(* INIT DIGITAL OUTPUT STUFF *)
FB_DO_SW_001.InitMqtt(MQTTPublishPrefix:= ADR(MqttPubSwitchPrefix),					(* pointer to string prefix for the mqtt publish topic *)
	MQTTSubscribePrefix:= ADR(MqttSubSwitchPrefix),									(* pointer to string prefix for the mqtt subscribe topic *)
	pMqttPublishQueue := ADR(MqttVariables.fbMqttPublishQueue),						(* pointer to MqttPublishQueue to send a new Mqtt event *)
	pMqttCallbackCollector := ADR(MqttVariables.collector_FB_OUTPUT_SWITCH_MQTT)	(* pointer to CallbackCollector to receive Mqtt subscription events *)
);
FB_DO_SW_002.InitMqtt(MQTTPublishPrefix:= ADR(MqttPubSwitchPrefix),	MQTTSubscribePrefix:= ADR(MqttSubSwitchPrefix), pMqttPublishQueue := ADR(MqttVariables.fbMqttPublishQueue), pMqttCallbackCollector := ADR(MqttVariables.collector_FB_OUTPUT_SWITCH_MQTT));
FB_DO_SW_003.InitMqtt(MQTTPublishPrefix:= ADR(MqttPubSwitchPrefix),	MQTTSubscribePrefix:= ADR(MqttSubSwitchPrefix),	pMqttPublishQueue := ADR(MqttVariables.fbMqttPublishQueue), pMqttCallbackCollector := ADR(MqttVariables.collector_FB_OUTPUT_SWITCH_MQTT));
FB_DO_SW_004.InitMqtt(MQTTPublishPrefix:= ADR(MqttPubSwitchPrefix),	MQTTSubscribePrefix:= ADR(MqttSubSwitchPrefix),	pMqttPublishQueue := ADR(MqttVariables.fbMqttPublishQueue), pMqttCallbackCollector := ADR(MqttVariables.collector_FB_OUTPUT_SWITCH_MQTT));
FB_DO_SW_005.InitMqtt(MQTTPublishPrefix:= ADR(MqttPubSwitchPrefix),	MQTTSubscribePrefix:= ADR(MqttSubSwitchPrefix),	pMqttPublishQueue := ADR(MqttVariables.fbMqttPublishQueue), pMqttCallbackCollector := ADR(MqttVariables.collector_FB_OUTPUT_SWITCH_MQTT));
FB_DO_SW_006.InitMqtt(MQTTPublishPrefix:= ADR(MqttPubSwitchPrefix),	MQTTSubscribePrefix:= ADR(MqttSubSwitchPrefix),	pMqttPublishQueue := ADR(MqttVariables.fbMqttPublishQueue), pMqttCallbackCollector := ADR(MqttVariables.collector_FB_OUTPUT_SWITCH_MQTT));
FB_DO_SW_007.InitMqtt(MQTTPublishPrefix:= ADR(MqttPubSwitchPrefix),	MQTTSubscribePrefix:= ADR(MqttSubSwitchPrefix),	pMqttPublishQueue := ADR(MqttVariables.fbMqttPublishQueue), pMqttCallbackCollector := ADR(MqttVariables.collector_FB_OUTPUT_SWITCH_MQTT));
FB_DO_SW_008.InitMqtt(MQTTPublishPrefix:= ADR(MqttPubSwitchPrefix),	MQTTSubscribePrefix:= ADR(MqttSubSwitchPrefix),	pMqttPublishQueue := ADR(MqttVariables.fbMqttPublishQueue), pMqttCallbackCollector := ADR(MqttVariables.collector_FB_OUTPUT_SWITCH_MQTT));
FB_DO_SW_009.InitMqtt(MQTTPublishPrefix:= ADR(MqttPubSwitchPrefix),	MQTTSubscribePrefix:= ADR(MqttSubSwitchPrefix),	pMqttPublishQueue := ADR(MqttVariables.fbMqttPublishQueue), pMqttCallbackCollector := ADR(MqttVariables.collector_FB_OUTPUT_SWITCH_MQTT));
FB_DO_SW_010.InitMqtt(MQTTPublishPrefix:= ADR(MqttPubSwitchPrefix),	MQTTSubscribePrefix:= ADR(MqttSubSwitchPrefix),	pMqttPublishQueue := ADR(MqttVariables.fbMqttPublishQueue), pMqttCallbackCollector := ADR(MqttVariables.collector_FB_OUTPUT_SWITCH_MQTT));
FB_DO_SW_011.InitMqtt(MQTTPublishPrefix:= ADR(MqttPubSwitchPrefix),	MQTTSubscribePrefix:= ADR(MqttSubSwitchPrefix),	pMqttPublishQueue := ADR(MqttVariables.fbMqttPublishQueue), pMqttCallbackCollector := ADR(MqttVariables.collector_FB_OUTPUT_SWITCH_MQTT));
FB_DO_SW_012.InitMqtt(MQTTPublishPrefix:= ADR(MqttPubSwitchPrefix),	MQTTSubscribePrefix:= ADR(MqttSubSwitchPrefix), pMqttPublishQueue := ADR(MqttVariables.fbMqttPublishQueue), pMqttCallbackCollector := ADR(MqttVariables.collector_FB_OUTPUT_SWITCH_MQTT));
FB_DO_SW_013.InitMqtt(MQTTPublishPrefix:= ADR(MqttPubSwitchPrefix),	MQTTSubscribePrefix:= ADR(MqttSubSwitchPrefix), pMqttPublishQueue := ADR(MqttVariables.fbMqttPublishQueue), pMqttCallbackCollector := ADR(MqttVariables.collector_FB_OUTPUT_SWITCH_MQTT));
FB_DO_SW_014.InitMqtt(MQTTPublishPrefix:= ADR(MqttPubSwitchPrefix),	MQTTSubscribePrefix:= ADR(MqttSubSwitchPrefix), pMqttPublishQueue := ADR(MqttVariables.fbMqttPublishQueue), pMqttCallbackCollector := ADR(MqttVariables.collector_FB_OUTPUT_SWITCH_MQTT));
FB_DO_SW_015.InitMqtt(MQTTPublishPrefix:= ADR(MqttPubSwitchPrefix),	MQTTSubscribePrefix:= ADR(MqttSubSwitchPrefix), pMqttPublishQueue := ADR(MqttVariables.fbMqttPublishQueue), pMqttCallbackCollector := ADR(MqttVariables.collector_FB_OUTPUT_SWITCH_MQTT));
FB_DO_SW_016.InitMqtt(MQTTPublishPrefix:= ADR(MqttPubSwitchPrefix),	MQTTSubscribePrefix:= ADR(MqttSubSwitchPrefix), pMqttPublishQueue := ADR(MqttVariables.fbMqttPublishQueue), pMqttCallbackCollector := ADR(MqttVariables.collector_FB_OUTPUT_SWITCH_MQTT));
FB_DO_SW_017.InitMqtt(MQTTPublishPrefix:= ADR(MqttPubSwitchPrefix),	MQTTSubscribePrefix:= ADR(MqttSubSwitchPrefix), pMqttPublishQueue := ADR(MqttVariables.fbMqttPublishQueue), pMqttCallbackCollector := ADR(MqttVariables.collector_FB_OUTPUT_SWITCH_MQTT));
FB_DO_SW_018.InitMqtt(MQTTPublishPrefix:= ADR(MqttPubSwitchPrefix),	MQTTSubscribePrefix:= ADR(MqttSubSwitchPrefix), pMqttPublishQueue := ADR(MqttVariables.fbMqttPublishQueue), pMqttCallbackCollector := ADR(MqttVariables.collector_FB_OUTPUT_SWITCH_MQTT));
FB_DO_SW_019.InitMqtt(MQTTPublishPrefix:= ADR(MqttPubSwitchPrefix),	MQTTSubscribePrefix:= ADR(MqttSubSwitchPrefix), pMqttPublishQueue := ADR(MqttVariables.fbMqttPublishQueue), pMqttCallbackCollector := ADR(MqttVariables.collector_FB_OUTPUT_SWITCH_MQTT));
FB_DO_SW_020.InitMqtt(MQTTPublishPrefix:= ADR(MqttPubSwitchPrefix),	MQTTSubscribePrefix:= ADR(MqttSubSwitchPrefix), pMqttPublishQueue := ADR(MqttVariables.fbMqttPublishQueue), pMqttCallbackCollector := ADR(MqttVariables.collector_FB_OUTPUT_SWITCH_MQTT));
FB_DO_SW_021.InitMqtt(MQTTPublishPrefix:= ADR(MqttPubSwitchPrefix),	MQTTSubscribePrefix:= ADR(MqttSubSwitchPrefix), pMqttPublishQueue := ADR(MqttVariables.fbMqttPublishQueue), pMqttCallbackCollector := ADR(MqttVariables.collector_FB_OUTPUT_SWITCH_MQTT));
FB_DO_SW_022.InitMqtt(MQTTPublishPrefix:= ADR(MqttPubSwitchPrefix),	MQTTSubscribePrefix:= ADR(MqttSubSwitchPrefix), pMqttPublishQueue := ADR(MqttVariables.fbMqttPublishQueue), pMqttCallbackCollector := ADR(MqttVariables.collector_FB_OUTPUT_SWITCH_MQTT));
FB_DO_SW_023.InitMqtt(MQTTPublishPrefix:= ADR(MqttPubSwitchPrefix),	MQTTSubscribePrefix:= ADR(MqttSubSwitchPrefix), pMqttPublishQueue := ADR(MqttVariables.fbMqttPublishQueue), pMqttCallbackCollector := ADR(MqttVariables.collector_FB_OUTPUT_SWITCH_MQTT));
FB_DO_SW_024.InitMqtt(MQTTPublishPrefix:= ADR(MqttPubSwitchPrefix),	MQTTSubscribePrefix:= ADR(MqttSubSwitchPrefix), pMqttPublishQueue := ADR(MqttVariables.fbMqttPublishQueue), pMqttCallbackCollector := ADR(MqttVariables.collector_FB_OUTPUT_SWITCH_MQTT));
FB_DO_SW_025.InitMqtt(MQTTPublishPrefix:= ADR(MqttPubSwitchPrefix),	MQTTSubscribePrefix:= ADR(MqttSubSwitchPrefix), pMqttPublishQueue := ADR(MqttVariables.fbMqttPublishQueue), pMqttCallbackCollector := ADR(MqttVariables.collector_FB_OUTPUT_SWITCH_MQTT));
FB_DO_SW_026.InitMqtt(MQTTPublishPrefix:= ADR(MqttPubSwitchPrefix),	MQTTSubscribePrefix:= ADR(MqttSubSwitchPrefix), pMqttPublishQueue := ADR(MqttVariables.fbMqttPublishQueue), pMqttCallbackCollector := ADR(MqttVariables.collector_FB_OUTPUT_SWITCH_MQTT));
FB_DO_SW_027.InitMqtt(MQTTPublishPrefix:= ADR(MqttPubSwitchPrefix),	MQTTSubscribePrefix:= ADR(MqttSubSwitchPrefix), pMqttPublishQueue := ADR(MqttVariables.fbMqttPublishQueue), pMqttCallbackCollector := ADR(MqttVariables.collector_FB_OUTPUT_SWITCH_MQTT));
FB_DO_SW_028.InitMqtt(MQTTPublishPrefix:= ADR(MqttPubSwitchPrefix),	MQTTSubscribePrefix:= ADR(MqttSubSwitchPrefix), pMqttPublishQueue := ADR(MqttVariables.fbMqttPublishQueue), pMqttCallbackCollector := ADR(MqttVariables.collector_FB_OUTPUT_SWITCH_MQTT));
FB_DO_SW_029.InitMqtt(MQTTPublishPrefix:= ADR(MqttPubSwitchPrefix),	MQTTSubscribePrefix:= ADR(MqttSubSwitchPrefix), pMqttPublishQueue := ADR(MqttVariables.fbMqttPublishQueue), pMqttCallbackCollector := ADR(MqttVariables.collector_FB_OUTPUT_SWITCH_MQTT));
FB_DO_SW_030.InitMqtt(MQTTPublishPrefix:= ADR(MqttPubSwitchPrefix),	MQTTSubscribePrefix:= ADR(MqttSubSwitchPrefix), pMqttPublishQueue := ADR(MqttVariables.fbMqttPublishQueue), pMqttCallbackCollector := ADR(MqttVariables.collector_FB_OUTPUT_SWITCH_MQTT));

(* INIT COVERS STUFF *)
FB_DO_COVER_001.InitMqtt(MQTTPublishPrefix:= ADR(MqttPubCoverPrefix),				(* pointer to string prefix for the mqtt publish topic *)
	MQTTSubscribePrefix:= ADR(MqttSubCoverPrefix),									(* pointer to string prefix for the mqtt subscribe topic *)
	pMqttPublishQueue := ADR(MqttVariables.fbMqttPublishQueue),						(* pointer to MqttPublishQueue to send a new Mqtt event *)
	pMqttCallbackCollector := ADR(MqttVariables.collector_FB_OUTPUT_COVER_MQTT), 	(* pointer to CallbackCollector to receive Mqtt subscription events *)
	MQTT.QoS.ExactlyOnce, 														(* specify the QoS for the POS mqtt events (values 0-100) *)
	2																				(* specify the resolution for the POS mqtt events *)
);

FB_DO_COVER_001.ConfigureFunctionBlock(T_LOCKOUT:=T#1S,								(* delay between change of direction *)
	T_UD:=T#20S																		(* run time to move the cover completely up/down *)
);

(* INIT VIRTUAL STUFF *)
FB_VIRTUAL_STRING_001.InitMqtt(MQTTPublishPrefix:= ADR(MqttPubVirtualPrefix),				
	MQTTSubscribePrefix:= ADR(MqttSubVirtualPrefix),									
	pMqttPublishQueue := ADR(MqttVariables.fbMqttPublishQueue),						
	pMqttCallbackCollector := ADR(MqttVariables.collector_FB_VIRTUAL_MQTT),
	MqttQos:=MQTT.QoS.ExactlyOnce, 
	MqttRetain:=FALSE									
);
FB_VIRTUAL_STRING_001.ConfigureFunctionBlockAsVirtualInput(DefaultValue:='HelloWorld',SetDefaultValueStartup:=TRUE,PublishAtStartup:=TRUE,UsePersistentAtStartup:=FALSE,ConfirmReceival:=TRUE);


FB_VIRTUAL_INT_001.InitMqtt(MQTTPublishPrefix:= ADR(MqttPubVirtualPrefix),				
	MQTTSubscribePrefix:= ADR(MqttSubVirtualPrefix),									
	pMqttPublishQueue := ADR(MqttVariables.fbMqttPublishQueue),						
	pMqttCallbackCollector := ADR(MqttVariables.collector_FB_VIRTUAL_MQTT),
	MqttQos:=MQTT.QoS.ExactlyOnce, 
	MqttRetain:=FALSE												
);
FB_VIRTUAL_INT_001.ConfigureFunctionBlockAsVirtualInput(DefaultValue:=0,SetDefaultValueStartup:=TRUE,PublishAtStartup:=TRUE,UsePersistentAtStartup:=FALSE,ConfirmReceival:=TRUE);
(* FB_VIRTUAL_INT_001.ConfigureFunctionBlockAsVirtualOutput(PublishAtStartup:=TRUE); *)


FB_VIRTUAL_BOOL_001.InitMqtt(MQTTPublishPrefix:= ADR(MqttPubVirtualPrefix),				
	MQTTSubscribePrefix:= ADR(MqttSubVirtualPrefix),									
	pMqttPublishQueue := ADR(MqttVariables.fbMqttPublishQueue),						
	pMqttCallbackCollector := ADR(MqttVariables.collector_FB_VIRTUAL_MQTT),
	MqttQos:=MQTT.QoS.ExactlyOnce, 
	MqttRetain:=FALSE											
);
(* FB_VIRTUAL_BOOL_001.ConfigureFunctionBlockAsVirtualInput(DefaultValue:=FALSE,SetDefaultValueStartup:=TRUE,PublishAtStartup:=TRUE,UsePersistentAtStartup:=FALSE); *)
FB_VIRTUAL_BOOL_001.ConfigureFunctionBlockAsVirtualOutput(PublishAtStartup:=TRUE);

FB_VIRTUAL_REAL_001.InitMqtt(MQTTPublishPrefix:= ADR(MqttPubVirtualPrefix),				
	MQTTSubscribePrefix:= ADR(MqttSubVirtualPrefix),									
	pMqttPublishQueue := ADR(MqttVariables.fbMqttPublishQueue),						
	pMqttCallbackCollector := ADR(MqttVariables.collector_FB_VIRTUAL_MQTT),
	MqttQos:=MQTT.QoS.ExactlyOnce, 
	MqttRetain:=FALSE												
);
FB_VIRTUAL_REAL_001.ConfigureFunctionBlockAsVirtualInput(DefaultValue:=0.1,SetDefaultValueStartup:=TRUE,PublishAtStartup:=TRUE,UsePersistentAtStartup:=FALSE,ConfirmReceival:=TRUE);
(* FB_VIRTUAL_REAL_001.ConfigureFunctionBlockAsVirtualOutput(PublishAtStartup:=TRUE); *)


(* INIT BISTABLE RELAIS *) 
FB_DO_BISTABLE_001.InitMqtt(MQTTPublishPrefix:= ADR(MqttPubSwitchPrefix),	MQTTSubscribePrefix:= ADR(MqttSubSwitchPrefix), pMqttPublishQueue := ADR(MqttVariables.fbMqttPublishQueue), pMqttCallbackCollector := ADR(MqttVariables.collector_FB_OUTPUT_SWITCH_MQTT));
FB_DO_BISTABLE_001.ConfigureFunctionBlock(T_hold:=T#10S); 

                    
END_ACTION

ACTION MOVE_COVERS:
                      FB_DO_COVER_001(
	UP:=FB_DI_PB_013.P_LONG,
	DN:=FB_DI_PB_015.P_LONG,
	MU=>DO_031,
	MD=>DO_032	
	);
                    
END_ACTION

ACTION PROCESS_VIRTUAL:
                      
FB_VIRTUAL_BOOL_001();
FB_VIRTUAL_INT_001();
FB_VIRTUAL_STRING_001();
FB_VIRTUAL_REAL_001();
                    
END_ACTION
END_PROGRAM

PROGRAM PLC_PRG_MQTT
  VAR
    broker : STRING := '192.168.1.52:1883';  (* variables for MQTT configuration *)
    clientID : STRING := 'PLC-House';  (* use the below for username password authentication to broker broker :STRING:='user:password@192.168.1.36:1883'; user led to indicate broker status, é!COCKPIT version LED_1_BrokerStatus :FbAppLED; *)
    MQTTClient : MQTT.MQTTClient;
    MQTT_IN_OUT : MQTT.MQTT_IN_OUT;
    MQTTInfo : MQTT.MQTT_INFO;
    MQTTLwtTopic : STRING := 'Devices/PLC/House/availability';
    MQTTLwtPayload : STRING := 'offline';
    MQTTBirthMessage : MQTT_MESSAGE;
    MQTTBirthTopic : STRING := 'Devices/PLC/House/availability';
    MQTTBirthPayload : STRING := 'online';
    MQTTBirthHartbeat : OSCAT_BASIC.GEN_PULSE;
    MQTTBirthHartbeatTime : TIME := TIME#5s0ms;
    MQTTConnectTrigger : Standard.R_TRIG;
    MQTTPublishBirth : BOOL := TRUE;
    MQTTBirthPublisher : FB_MqttPublishWorker;
    initMqtt : BOOL;  (* variables for MQTT setup *)
    icounter : UDINT;
    ipublishers : UDINT := 40;  (* variables for MQTT publishing *)
    publishers : ARRAY[0..39] OF FB_MqttPublishWorker;
    i : UDINT;  (* variables to work with Mqttbuffer *)
    subscriber_FB_OUTPUT_SWITCH_MQTT : MQTT.MQTTSubscribe;  (* variables for MQTT subscribing *)
    subscriber_FB_OUTPUT_COVER_MQTT : MQTT.MQTTSubscribe;
    subscriber_FB_VIRTUAL_MQTT : MQTT.MQTTSubscribe;
    subscriber_FB_DIMMER_MQTT : MQTT.MQTTSubscribe;
  END_VAR

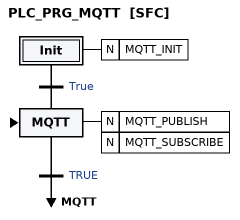
INITIAL_STEP Init:
  MQTT_INIT(N);
END_STEP
TRANSITION FROM Init TO MQTT
  := True;
END_TRANSITION
STEP MQTT:
  MQTT_PUBLISH(N);
  MQTT_SUBSCRIBE(N);
END_STEP
TRANSITION FROM MQTT TO MQTT
  := TRUE;
END_TRANSITION

ACTION MQTT_INIT:
                      
IF NOT initMqtt THEN
	initMqtt := TRUE;
	(* Basic MQTT config *)
	MQTT_IN_OUT.ClientID := clientID;
	
	(* Set the LWT topic / payload *)
	MQTT_IN_OUT.BuildWillTopicAndMessage := FALSE;
	MQTT_IN_OUT.WillTopicBase := '';
	MQTT_IN_OUT.ClientWillTopic := MQTTLwtTopic;
	MQTT_IN_OUT.ClientWillMessage := MQTTLwtPayload;
	
	(* Set the birth message *)
	MQTTBirthMessage.Payload := MQTTBirthPayload;
	MQTTBirthMessage.Topic := MQTTBirthTopic;
	MQTTBirthMessage.Qos := MqttVariables.MQTT_QOS_EXACTLY_ONCE;
	MQTTBirthMessage.MqttRetain := FALSE;
	
	(* Configure the rising edge detector to detect a connect/reconnect to the broker, used for  birth message *)
	MQTTConnectTrigger(CLK := MQTTInfo.MQTT_CONNECTED);
	
	(* Configure the dedicated MQTTBirth publisher *)
	MQTTBirthPublisher.Init(inputMQTT_IN_OUT:= ADR(MQTT_IN_OUT));
	
	(* Configure the pulse generator for the birth message hartbeat *)
	 MQTTBirthHartbeat(ENQ:=TRUE, PTH:=T#0S, PTL:=MQTTBirthHartbeatTime);
	
	(* INIT MQTT PUBLISH STUFF *)
	FOR icounter := 0 TO (ipublishers-1) DO		
		publishers[icounter].Init(inputMQTT_IN_OUT:= ADR(MQTT_IN_OUT));
	END_FOR 
	
	(* INIT MQTT SUBSCRIBE STUFF *)
	subscriber_FB_OUTPUT_SWITCH_MQTT.SetMqttInOut(MQTT_IN_OUT:= MQTT_IN_OUT);	
	subscriber_FB_OUTPUT_COVER_MQTT.SetMqttInOut(MQTT_IN_OUT:= MQTT_IN_OUT);
	subscriber_FB_VIRTUAL_MQTT.SetMqttInOut(MQTT_IN_OUT:= MQTT_IN_OUT);	
	subscriber_FB_DIMMER_MQTT.SetMqttInOut(MQTT_IN_OUT:= MQTT_IN_OUT);

END_IF


                    
END_ACTION

ACTION MQTT_PUBLISH:
                      (* set user led green if connected to MQTT broker, flashing red if not *)
(* é!COCKPIT version *)
(* LED_1_BrokerStatus(eID:=eLedID.AppLED_1, xOpen:=TRUE );
IF(MQTTClient.connected) THEN
	LED_1_BrokerStatus.SetStatic(eLedColor.Green);
ELSE
	LED_1_BrokerStatus.SetFlash(T#1S,eLedColor.Red, eLedColor.Off);  
END_IF *)
(* Codesys 3S version *)
(*
IF MQTTClient.connected THEN
     PFC.SetLed(which:=PFC.LED.U1, how:=PFC.LedState.STATIC_GRN);
ELSE
     PFC.SetLed(which:=PFC.LED.U1, how:=PFC.LedState.BLINK_RED);
END_IF 
*)

(* allow the rising edge detector to detect a connect/reconnect to the broker, used for  birth message *)
MQTTConnectTrigger(CLK := MQTTInfo.MQTT_CONNECTED);

(* allow the pulse generator to generate a pulse, used for birth message hartbeat *)
MQTTBirthHartbeat(ENQ:=TRUE, PTH:=T#0S, PTL:=MQTTBirthHartbeatTime);

(* Check if this is a new connection due to startup or connection issues *)
IF initMqtt AND (MQTTConnectTrigger.Q OR MQTTBirthHartbeat.Q) THEN
	MQTTPublishBirth := TRUE;
END_IF

(* On connect or reconnect publish a birth message using the dedicated birth publisher *)
IF MQTTPublishBirth THEN
	MQTTBirthPublisher.PublishMessage(MqttMessage := MQTTBirthMessage);
	MQTTPublishBirth:=FALSE;
END_IF


(* Check if Mqtt is initialized AND if there are elements on the queue to process AND if a MQTTbirthmessage has been published successfully *)
IF initMqtt AND NOT(MqttVariables.fbMqttPublishQueue.EMPTY) AND MQTTPublishBirth = FALSE AND MQTTBirthPublisher.SendDone THEN	
	(* Loop through all free publishers untill there are no more elements in the queue or no more free publishers *)
	FOR i:=0 TO (ipublishers-1) DO			
		(* use the publishers that are free  *)
		IF publishers[i].SendDone AND NOT(MqttVariables.fbMqttPublishQueue.EMPTY) THEN	
			(* Pass message from the queue to a publisher *)
			publishers[i].PublishMessage(MqttMessage:= MqttVariables.fbMqttPublishQueue.GetMessage());
		ELSIF MqttVariables.fbMqttPublishQueue.EMPTY THEN
			(* Queue is empty, jump out of the for loop	*)
			EXIT;	
		END_IF
	END_FOR
END_IF


(* If MQTT is initialized, let the MqttPublishWorkers do their work *)
IF initMqtt THEN	
	MQTT_IN_OUT.clientFB(
		MQTT_IN_OUT:= MQTT_IN_OUT, 
		ENABLE:= TRUE, 
		URL:= broker, 
		TIMEOUT:= T#1S, 
		TLS:= FALSE);		
		
	MQTTBirthPublisher();
	
	FOR i := 0 TO (ipublishers-1) DO
  		publishers[i]();
	END_FOR

END_IF

                    
END_ACTION

ACTION MQTT_SUBSCRIBE:
                      (* If MQTT is initialized, let the subscriber(s) do its work *)
IF initMqtt THEN
	
	MQTT_IN_OUT.clientFB(
		MQTT_IN_OUT:= MQTT_IN_OUT, 
		ENABLE:= TRUE, 
		URL:= broker, 
		TIMEOUT:= T#1S, 
		TLS:= FALSE);

	subscriber_FB_OUTPUT_SWITCH_MQTT(
		Subscribe:= TRUE, 
		Topic:= ADR('Devices/PLC/House/In/DigitalOutputs/+'), 
		QoSSubscribe:= MqttVariables.MQTT_QOS_EXACTLY_ONCE, 
		ExpectingString:= TRUE, 
		Callback:= MqttVariables.collector_FB_OUTPUT_SWITCH_MQTT,
	);
	
	subscriber_FB_OUTPUT_COVER_MQTT(
		Subscribe:= TRUE, 
		Topic:= ADR('Devices/PLC/House/In/Covers/+'), 
		QoSSubscribe:= MqttVariables.MQTT_QOS_EXACTLY_ONCE, 
		ExpectingString:= TRUE, 
		Callback:= MqttVariables.collector_FB_OUTPUT_COVER_MQTT,
	);
	
	subscriber_FB_VIRTUAL_MQTT(
		Subscribe:= TRUE, 
		Topic:= ADR('Devices/PLC/House/In/Virtuals/+'), 
		QoSSubscribe:= MqttVariables.MQTT_QOS_EXACTLY_ONCE, 
		ExpectingString:= TRUE, 
		Callback:= MqttVariables.collector_FB_VIRTUAL_MQTT,
	);
	subscriber_FB_DIMMER_MQTT(
		Subscribe:= TRUE, 
		Topic:= ADR('Devices/PLC/House/In/Dimmers/+'), 
		QoSSubscribe:= MqttVariables.MQTT_QOS_EXACTLY_ONCE, 
		ExpectingString:= TRUE, 
		Callback:= MqttVariables.collector_FB_DIMMER_MQTT,
	);
END_IF

                    
END_ACTION
END_PROGRAM

PROGRAM PLC_PRG_RS485
  VAR
    ModbusMaster : WagoAppPlcModbus.FbMbMasterSerial := (xConnect := TRUE, udiBaudrate := 9600, usiDataBits := 8, eParity := WagoTypesCom.eTTYParity.None, eStopBits := WagoTypesCom.eTTYStopBits.One, eHandshake := WagoTypesCom.eTTYHandshake.None, ePhysical := WagoTypesCom.eTTYPhysicalLayer.RS485_HalfDuplex, eFrameType := eMbFrameType.RTU, tTimeOut := TIME#500ms);  (* CODESYS 3S Version version xComPortOpen : BOOL; xComPortError : BOOL; rtsResult : RTS_IEC_RESULT; stComPortSettings : SysCom.SysComSettings :=( ulBaudrate :=9600, byParity := 0, byStopBits:=1, ulTimeout :=500, ulBufferSize :=256, sPort:=SYS_COM_PORTS.SYS_COMPORT1 ); hComPort : RTS_IEC_HANDLE; awReadBuffer : ARRAY[0..124] OF WORD; awWriteBuffer : ARRAY[0..124] OF WORD; fbModbusRequest : IoDrvModbus.ModbusRequest2; eComError : IoDrvModbus.MB_ErrorCodes; é!COCKPIT version *)
    RtuQuery : WagoAppPlcModbus.typMbQuery;
    RtuResponse : WagoAppPlcModbus.typMbResponse;
    Trigger : BOOL := FALSE;  (* Shared variables for é!COCKPIT and CODESYS 3S Version *)
    InitRS485 : BOOL := FALSE;
    ActiveRtuQuery : RS485_RtuQuery;
    RS485BusController : FB_RS485_BUSCONTROLLER;
    MqttRS485Prefix : STRING(100) := 'Devices/PLC/House/Out/RS485/';  (* RS485 *)
    FB_RS485_EASTRON_SDM220_1 : FB_RS485_EASTRON_SDM220_MQTT;
    FB_RS485_ESERA_1WIRE_GATEWAY_MQTT_HOME : FB_RS485_ESERA_1WIRE_GATEWAY_MQTT;
  END_VAR

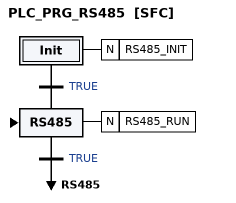
INITIAL_STEP Init:
  RS485_INIT(N);
END_STEP
TRANSITION FROM Init TO RS485
  := TRUE;
END_TRANSITION
STEP RS485:
  RS485_RUN(N);
END_STEP
TRANSITION FROM RS485 TO RS485
  := TRUE;
END_TRANSITION

ACTION RS485_RUN:
                      (* CODESYS 3S Version version*)
(*
IF(NOT xComPortOpen AND NOT xComPortError) THEN
    hComPort := SysCom.SysComOpen2( pSettings := ADR(stComPortSettings), pSettingsEx := 0, pResult := ADR(rtsResult));     
    xComPortError := (hComPort = RTS_INVALID_HANDLE OR rtsResult <> 0);
    xComPortOpen := NOT xComPortError;
END_IF


IF xComPortOpen THEN
	fbModbusRequest.modbusCommand.uiFunctionCode := RS485BusController.ActiveRtuQuery.FunctionCode;
    fbModbusRequest.modbusCommand.uiReadOffset := RS485BusController.ActiveRtuQuery.ReadAddress;	
    fbModbusRequest.modbusCommand.uiReadLen :=RS485BusController.ActiveRtuQuery.ReadQuantity;	   
    fbModbusRequest.pRecvData := ADR(awReadBuffer);
    fbModbusRequest.pSendData := ADR(awWriteBuffer);        
    fbModbusRequest.tResponseTimeout := T#1S;
	fbModbusRequest.transmission := MB_Transmission.RTU;
    fbModbusRequest(
        hComPort := hComPort,
        xExecute := Trigger,
        usiSlaveAddr := RS485BusController.ActiveRtuQuery.DeviceId,		
        byModbusError => eComError);
		
END_IF
*)
	
(* é!COCKPIT version*)
RtuQuery.bUnitId := RS485BusController.ActiveRtuQuery.DeviceId;	
RtuQuery.bFunctionCode := RS485BusController.ActiveRtuQuery.FunctionCode;	
RtuQuery.uiReadAddress := RS485BusController.ActiveRtuQuery.ReadAddress;	
RtuQuery.uiReadQuantity := RS485BusController.ActiveRtuQuery.ReadQuantity;
ModbusMaster(
	I_Port := IoConfig_Globals.COM1,
	utQuery:= RtuQuery,
	xTrigger := Trigger,
	utResponse:= RtuResponse);


(* Shared variables for é!COCKPIT and CODESYS 3S Version *)
RS485BusController();

(* RS485 devices *)
FB_RS485_EASTRON_SDM220_1();
FB_RS485_ESERA_1WIRE_GATEWAY_MQTT_HOME();
                    
END_ACTION

ACTION RS485_INIT:
                      IF NOT InitRS485 THEN
	InitRS485 := TRUE;

(* INIT RS485 BUS CONTROLLER; CODESYS 3S Version version *)
(*
RS485BusController.Init(
	StartupDelay := T#5S,				(* Time to wait after startup to start using the bus, prevents boot delay issues when RS485 are not ready yet on startup *)		
	SilenceTime := T#50MS,				(* Silence time between two requests, important to not get faulty data on bus *)
	BusTrigger := ADR(Trigger),			(* Pointer to the bool used to initiate bus requests *)
	BusData := ADR(awReadBuffer),		(* Pointer to the array containing the bus response data *)
	BusError := ADR(xComPortError)		(* Pointer to the bus error bool *)
);
*)

(* INIT RS485 BUS CONTROLLER; é!COCKPIT version *)
RS485BusController.Init(
	StartupDelay := T#5S,				(* Time to wait after startup to start using the bus, prevents boot delay issues when RS485 are not ready yet on startup *)		
	SilenceTime := T#50MS,				(* Silence time between two requests, important to not get faulty data on bus *)
	BusTrigger := ADR(Trigger),			(* Pointer to the bool used to initiate bus requests *)
	BusData := ADR(RtuResponse.awData),	(* Pointer to the array containing the bus response data *)
	BusError := ADR(ModbusMaster.xError)(* Pointer to the bus error bool *)
);

RS485BusController.RegisterDevice(device := FB_RS485_EASTRON_SDM220_1);
RS485BusController.RegisterDevice(device := FB_RS485_ESERA_1WIRE_GATEWAY_MQTT_HOME);

(* INIT RS485 DEVICE STUFF *)
FB_RS485_EASTRON_SDM220_1.InitRS485(
	Data1PollingInterval := T#10S,		(* Polling interval for data array 1 *)				
	Data2PollingInterval := T#20S,		(* Polling interval for data array 2 *)			
	Data3PollingInterval := T#30S,		(* Polling interval for data array 3 *)			
	DeviceAddress := 1					(* Device address of the modbus device *)			
);

FB_RS485_EASTRON_SDM220_1.InitMqtt(
	MQTTPublishPrefix:= ADR(MqttRS485Prefix),						(* pointer to string prefix for the mqtt publish topic *)
	pMqttPublishQueue := ADR(MqttVariables.fbMqttPublishQueue)		(* pointer to MqttPublishQueue to send a new Mqtt event *)
);

FB_RS485_ESERA_1WIRE_GATEWAY_MQTT_HOME.InitRS485(
	DeviceAddress := 2
);

FB_RS485_ESERA_1WIRE_GATEWAY_MQTT_HOME.InitMqtt(
	MQTTPublishPrefix:= ADR(MqttRS485Prefix),	
	pMqttPublishQueue := ADR(MqttVariables.fbMqttPublishQueue)
);

(* ENABLE OWD DEVICES ON ESARE GATEWAY *)
FB_RS485_ESERA_1WIRE_GATEWAY_MQTT_HOME.EnableOwd(
	OwdNumber := 1,
	DataPollingInterval := T#2M
);

FB_RS485_ESERA_1WIRE_GATEWAY_MQTT_HOME.EnableOwd(
	OwdNumber := 2,
	DataPollingInterval := T#2M
);


END_IF
                    
END_ACTION
END_PROGRAM

CONFIGURATION Application
  RESOURCE HomeAutomation ON PLC
    {attribute 'qualified_only'}
    VAR_GLOBAL  (* MqttVariables *)
      fbMqttPublishQueue : FB_MqttPublishQueue;  (* Shared Variables for MQTT publish communication *)
      collector_FB_OUTPUT_SWITCH_MQTT : MQTT.CallbackCollector;  (* Shared Variables for MQTT subscribe communication *)
      collector_FB_OUTPUT_COVER_MQTT : MQTT.CallbackCollector;
      collector_FB_VIRTUAL_MQTT : MQTT.CallbackCollector;
      collector_FB_DIMMER_MQTT : MQTT.CallbackCollector;
      MQTT_QOS_EXACTLY_ONCE : MQTT.QoS := MQTT.QoS.ExactlyOnce;  (* QOS Constants *)
    END_VAR
    TASK MainTask(INTERVAL := T#50ms, PRIORITY := 4);
    TASK MqttCommunication(PRIORITY := 5);
    TASK RS485(INTERVAL := T#200ms, PRIORITY := 15);
    PROGRAM PLC_PRG_MAIN WITH MainTask : PLC_PRG_MAIN;
    PROGRAM PLC_PRG_MQTT WITH MqttCommunication : PLC_PRG_MQTT;
    PROGRAM PLC_PRG_RS485 WITH RS485 : PLC_PRG_RS485;
  END_RESOURCE
END_CONFIGURATION
